// TIA Portal V21 export
// export: Created 2026-11-11T00:47:19.1187632Z, ExportSetting WithDefaults, DisplayName Totally Integrated Automation Portal, DisplayVersion V21 Update 3, DisplayName STEP 7 Professional, DisplayVersion V21 Update 3, DisplayName STEP 7 Safety, DisplayVersion V21, DisplayName Tech WebApplication, DisplayVersion V21, DisplayName WinCC Basic/Comfort/Advanced, DisplayVersion V21 Update 3, DisplayName WinCC Unified, DisplayVersion V21 Update 3
FUNCTION_BLOCK "FB_Fbd_ex051"   // FB361, FBD
{ S7_Optimized_Access := 'TRUE' }
VERSION : 0.1
// stored: AutoNumber true, IsIECCheckEnabled false, IsRetainMemResEnabled false, MemoryReserve 100, SetENOAutomatically false, UDAEnableTagReadback false
   VAR_INPUT
      v_mode : Int;
      v_f_id : HW_IO;
      v_mlen : UInt;
   END_VAR
   VAR_OUTPUT
      v_new : Bool;
      v_status : DWord;
      v_id : HW_IO;
      v_len : UInt;
   END_VAR
   VAR_IN_OUT
      v_tinfo : Array[0..99] of Byte;
      v_ainfo : Array[0..99] of Byte;
   END_VAR
   VAR
      inst { S7_SetPoint := 'True'} : RALRM;
   END_VAR
BEGIN

REGION Network 1: Description RALRM
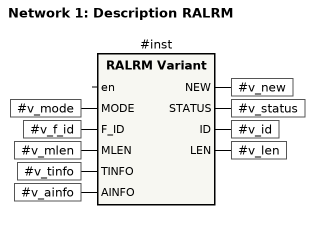
   #inst(MODE := #v_mode,   // RALRM
         F_ID := #v_f_id,
         MLEN := #v_mlen,
         TINFO := #v_tinfo,
         AINFO := #v_ainfo,
         NEW => #v_new,
         STATUS => #v_status,
         ID => #v_id,
         LEN => #v_len);
END_REGION
END_FUNCTION_BLOCK
